// TIA Portal V20 export
// export: Created 2026-10-09T07:03:58.1914004Z, ExportSetting WithDefaults, DisplayName Totally Integrated Automation Portal, DisplayVersion V20, DisplayName TIA Portal Openness, DisplayVersion V20, DisplayName TIA Portal Teamcenter Gateway, DisplayVersion V20, DisplayName TIA Portal Version Control Interface, DisplayVersion V20, DisplayName SINAMICS Startdrive Advanced, DisplayVersion V20 SP1 Update 2, DisplayName SINAMICS Startdrive G110M, G120, G120C, G120D, G120P, G115D, DisplayVersion V20 SP1 Update 2, DisplayName SINAMICS Startdrive G130, G150, S120, S150, SINAMICS MV, G220, S200, S210, DisplayVersion V20 SP1 Update 2, DisplayName STEP 7 Professional, DisplayVersion V20, DisplayName STEP 7 Safety, DisplayVersion V20, DisplayName WinCC Basic/Comfort/Advanced, DisplayVersion V20, DisplayName WinCC Professional, DisplayVersion V20, DisplayName WinCC Unified, DisplayVersion V20
FUNCTION_BLOCK "FB_GRAPH_PressDemoHome"   // FB100, GRAPH
VERSION : 0.1
// stored: AcknowledgeErrorsRequired true, AutoNumber true, GraphVersion 6.0, InitialValuesAcquisition false, IsIECCheckEnabled false, LanguageInNetworks LAD, LockOperatingMode false, PermanentILProcessingInMANMode false, SetENOAutomatically false, SkipSteps false, UDAEnableTagReadback false, WithAlarmHandling true
   // inherited from GRAPH_BASE
   VAR
      OFF_SQ_BASE : Bool;
   END_VAR
   VAR_INPUT
      OFF_SQ { ExternalAccessible := 'False'; ExternalVisible := 'False'; ExternalWritable := 'False'} : Bool := false;   // Turn sequence off
      INIT_SQ { ExternalAccessible := 'False'; ExternalVisible := 'False'; ExternalWritable := 'False'} : Bool := false;   // Set sequence to initial state
      ACK_EF { ExternalAccessible := 'False'; ExternalVisible := 'False'; ExternalWritable := 'False'} : Bool := false;   // Acknowledge all errors and faults
      S_PREV { ExternalAccessible := 'False'; ExternalVisible := 'False'; ExternalWritable := 'False'} : Bool := false;   // Output previous step in parameter S_NO
      S_NEXT { ExternalAccessible := 'False'; ExternalVisible := 'False'; ExternalWritable := 'False'} : Bool := false;   // Indicate next step in parameter S_NO
      SW_AUTO { ExternalAccessible := 'False'; ExternalVisible := 'False'; ExternalWritable := 'False'} : Bool := false;   // Automatic mode
      SW_TAP { ExternalAccessible := 'False'; ExternalVisible := 'False'; ExternalWritable := 'False'} : Bool := false;   // Semiautomatic/switch with transition
      SW_TOP { ExternalAccessible := 'False'; ExternalVisible := 'False'; ExternalWritable := 'False'} : Bool := false;   // Semiautomatic/ignore transition
      SW_MAN { ExternalAccessible := 'False'; ExternalVisible := 'False'; ExternalWritable := 'False'} : Bool := false;   // Manual mode
      S_SEL { ExternalAccessible := 'False'; ExternalVisible := 'False'; ExternalWritable := 'False'} : Int := 0;   // Select step to be output to S_NO
      S_ON { ExternalAccessible := 'False'; ExternalVisible := 'False'; ExternalWritable := 'False'} : Bool := false;   // Activate step indicated in S_NO
      S_OFF { ExternalAccessible := 'False'; ExternalVisible := 'False'; ExternalWritable := 'False'} : Bool := false;   // Disable step indicated in S_NO
      T_PUSH { ExternalAccessible := 'False'; ExternalVisible := 'False'; ExternalWritable := 'False'} : Bool := false;   // Enable transition to switch in semi automatic mode
      Run : BOOL;
      Reset : BOOL;
      OwnerIndex : DINT;
      Delta : TIME;
   END_VAR
   VAR_OUTPUT
      S_NO { ExternalAccessible := 'False'; ExternalVisible := 'False'; ExternalWritable := 'False'} : Int := 0;   // Step number
      S_MORE { ExternalAccessible := 'False'; ExternalVisible := 'False'; ExternalWritable := 'False'} : Bool := false;   // More steps are available and can be shown in S_NO
      S_ACTIVE { ExternalAccessible := 'False'; ExternalVisible := 'False'; ExternalWritable := 'False'} : Bool := false;   // Step indicated in S_NO is active
      ERR_FLT { ExternalAccessible := 'False'; ExternalVisible := 'False'; ExternalWritable := 'False'} : Bool := false;   // Interlock or supervision group error
      AUTO_ON { ExternalAccessible := 'False'; ExternalVisible := 'False'; ExternalWritable := 'False'} : Bool := false;   // Automatic mode is active
      TAP_ON { ExternalAccessible := 'False'; ExternalVisible := 'False'; ExternalWritable := 'False'} : Bool := false;   // Semiautomatic mode/step with transition enabled
      TOP_ON { ExternalAccessible := 'False'; ExternalVisible := 'False'; ExternalWritable := 'False'} : Bool := false;   // Semiautomatic mode/ignore transition enabled
      MAN_ON { ExternalAccessible := 'False'; ExternalVisible := 'False'; ExternalWritable := 'False'} : Bool := false;   // Manual mode is active
   END_VAR
   VAR_IN_OUT
      PressRam : "FB_CylinderCM";
      Door : "FB_CylinderCM";
      PartSlide : "FB_CylinderCM";
      Seq : "FRK_SequenceCtx";
      Row1 : "FRK_SequenceRow";
      Row2 : "FRK_SequenceRow";
      Row3 : "FRK_SequenceRow";
      Row4 : "FRK_SequenceRow";
      Ready1 { ExternalAccessible := 'False'; ExternalVisible := 'False'; ExternalWritable := 'False'} : BOOL;
      Ready2 { ExternalAccessible := 'False'; ExternalVisible := 'False'; ExternalWritable := 'False'} : BOOL;
      Ready3 { ExternalAccessible := 'False'; ExternalVisible := 'False'; ExternalWritable := 'False'} : BOOL;
      Ready4 { ExternalAccessible := 'False'; ExternalVisible := 'False'; ExternalWritable := 'False'} : BOOL;
      Ready5 { ExternalAccessible := 'False'; ExternalVisible := 'False'; ExternalWritable := 'False'} : BOOL;
   END_VAR
BEGIN
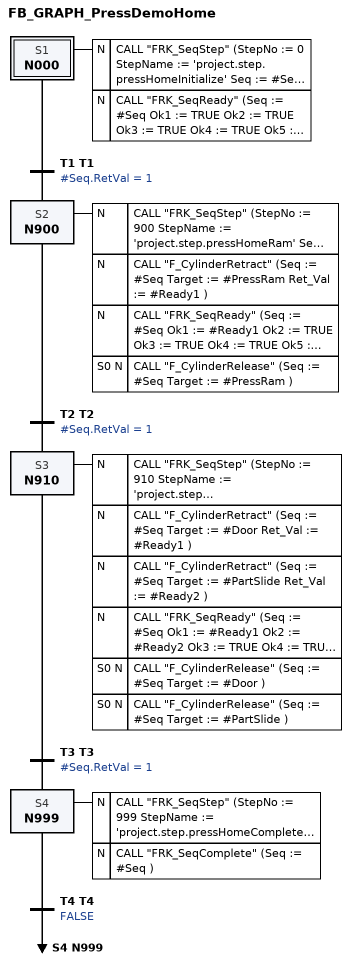
   // sequencer 1
   INITIAL_STEP N000:   // S1, max time T#10S, warning time T#7S
              N    CALL "FRK_SeqStep" 
                   (StepNo := 0
                   StepName := 'project.step.pressHomeInitialize'
                   Seq := #Seq
                   Row := #Row1
                   )
              N    CALL "FRK_SeqReady" 
                   (Seq := #Seq
                   Ok1 := TRUE
                   Ok2 := TRUE
                   Ok3 := TRUE
                   Ok4 := TRUE
                   Ok5 := TRUE
                   )
   END_STEP
   TRANSITION T1 FROM N000 TO N900   // T1
      := #Seq.RetVal = 1;
   END_TRANSITION
   STEP N900:   // S2, max time T#10S, warning time T#7S
              N    CALL "FRK_SeqStep" 
                   (StepNo := 900
                   StepName := 'project.step.pressHomeRam'
                   Seq := #Seq
                   Row := #Row2
                   )
              N    CALL "F_CylinderRetract" 
                   (Seq := #Seq
                   Target := #PressRam
                   Ret_Val := #Ready1
                   )
              N    CALL "FRK_SeqReady" 
                   (Seq := #Seq
                   Ok1 := #Ready1
                   Ok2 := TRUE
                   Ok3 := TRUE
                   Ok4 := TRUE
                   Ok5 := TRUE
                   )
          S0  N    CALL "F_CylinderRelease" 
                   (Seq := #Seq
                   Target := #PressRam
                   )
   END_STEP
   TRANSITION T2 FROM N900 TO N910   // T2
      := #Seq.RetVal = 1;
   END_TRANSITION
   STEP N910:   // S3, max time T#10S, warning time T#7S
              N    CALL "FRK_SeqStep" 
                   (StepNo := 910
                   StepName := 'project.step.pressHomeDoorAndSlide'
                   Seq := #Seq
                   Row := #Row3
                   )
              N    CALL "F_CylinderRetract" 
                   (Seq := #Seq
                   Target := #Door
                   Ret_Val := #Ready1
                   )
              N    CALL "F_CylinderRetract" 
                   (Seq := #Seq
                   Target := #PartSlide
                   Ret_Val := #Ready2
                   )
              N    CALL "FRK_SeqReady" 
                   (Seq := #Seq
                   Ok1 := #Ready1
                   Ok2 := #Ready2
                   Ok3 := TRUE
                   Ok4 := TRUE
                   Ok5 := TRUE
                   )
          S0  N    CALL "F_CylinderRelease" 
                   (Seq := #Seq
                   Target := #Door
                   )
          S0  N    CALL "F_CylinderRelease" 
                   (Seq := #Seq
                   Target := #PartSlide
                   )
   END_STEP
   TRANSITION T3 FROM N910 TO N999   // T3
      := #Seq.RetVal = 1;
   END_TRANSITION
   STEP N999:   // S4, max time T#10S, warning time T#7S
              N    CALL "FRK_SeqStep" 
                   (StepNo := 999
                   StepName := 'project.step.pressHomeComplete'
                   Seq := #Seq
                   Row := #Row4
                   )
              N    CALL "FRK_SeqComplete" 
                   (Seq := #Seq
                   )
   END_STEP
   TRANSITION T4 FROM N999 TO N999   // T4, jump
      := FALSE;
   END_TRANSITION
END_FUNCTION_BLOCK
